Fanuc KAREL source: ke00003.compact.KL

PROGRAM KE00003
%STACKSIZE=65535
%PRIORITY=65535
%NOLOCKGROUP
%ENVIRONMENT REGOPE
VAR
I : INTEGER
S : STRING[80]
STATUS : INTEGER
BEGIN
I=1
S='TEST'
SET_PREG_CMT(I,S,STATUS)
END KE00003
